FUNCTION FC 1 : VOID
BEGIN
NETWORK
      A I 0.0 @ home
END_FUNCTION
